(* IEC 61131-3 sources: CS_4_Aufzugsteuerung/src/Stations/CP112/Steuerung/Network, 1 file *)

(* ---- ConfigObjects.st ---- *)
FUNCTION GLOBAL TAB TASK_CONF
_K_TASK, _K_REAL,
_K_END_VAR,

_K_TASK, _K_CYCLIC,
_K_END_VAR,

_K_TASK, _K_BACKGROUND,
_K_END_VAR,

_K_END_CONF
END_FUNCTION

FUNCTION GLOBAL TAB IPR_CONF
_K_IPR
	0$UINT,
_K_END_VAR,
_K_END_CONF
END_FUNCTION

FUNCTION GLOBAL TAB CONFIG_TABLES
00096$UINT,
0$UINT, 1, 58, "_AXISBASE",
0$UINT, 1, 15, "_BUSINTERFACESDIASDRIVEMNG",
0$UINT, 0, 5, "_CAN",
0$UINT, 1, 11, "_CANLIB",
0$UINT, 1, 72, "_DRIVEAXIS",
0$UINT, 1, 81, "_DRIVEAXISBASE",
0$UINT, 1, 22, "_DRIVEAXISSET",
0$UINT, 1, 88, "_DRIVEMNG_DC062",
0$UINT, 1, 66, "_DRIVEMNGBASE",
0$UINT, 1, 20, "_FILESYS",
0$UINT, 0, 5, "_LINKER",
0$UINT, 1, 0, "_LMCABSENCODER",
0$UINT, 1, 117, "_LMCAXIS",
0$UINT, 2, 108, "_LMCAXISBASE",
0$UINT, 1, 32, "_LMCAXISREF",
0$UINT, 1, 41, "_LMCAXISVIS",
0$UINT, 1, 63, "_LMCAXISVISINT",
0$UINT, 1, 0, "_LMCAXISVISLOGHANDLE",
0$UINT, 1, 0, "_LMCAXISVISLOGVIEWER",
0$UINT, 1, 13, "_LMCAXISVISPARA",
0$UINT, 1, 1, "_LMCAXISVOVMONITORING",
0$UINT, 1, 75, "_LMCMATHFUNCTIONS",
0$UINT, 1, 1, "_LMCMODULEBASE",
0$UINT, 1, 0, "_LMCPUBLISHER",
0$UINT, 1, 11, "_LMCREFBASE",
0$UINT, 1, 21, "_LMCSAFETY",
0$UINT, 1, 1, "_MULTITASK",
0$UINT, 0, 5, "_OSKERNEL",
0$UINT, 1, 36, "_SERLIB",
0$UINT, 2, 0, "_STDLIB",
0$UINT, 1, 1, "_TASKOBJECTCONTROL",
0$UINT, 1, 69, "_VARANDRIVEBASE",
0$UINT, 1, 20, "AI043",
0$UINT, 1, 21, "ASCII_BIN",
0$UINT, 1, 26, "BUSINTERFACESDIAS",
0$UINT, 2, 1, "BUSINTERFACESDIASINTERNAL",
0$UINT, 1, 75, "BUSINTERFACEVARAN",
0$UINT, 0, 0, "CLSANTRIEB",
0$UINT, 0, 0, "CLSAUFZUGMODUL",
0$UINT, 0, 0, "CLSCOUNTER",
0$UINT, 0, 0, "CLSEMGSTOP_1",
0$UINT, 0, 0, "CLSENABLEDRIVE",
0$UINT, 0, 0, "CLSETAGENSENSORIK",
0$UINT, 0, 0, "CLSHAUPTABLAUF",
0$UINT, 0, 0, "CLSHMI",
0$UINT, 0, 0, "CLSMOTORCONTROL",
0$UINT, 0, 0, "CLSSIMPLECOUNTER",
0$UINT, 0, 0, "CLSTIMER",
0$UINT, 0, 0, "CLSTUERSENSORIK",
0$UINT, 1, 46, "CONTROLLER",
0$UINT, 1, 1, "CP112_IOS",
0$UINT, 0, 4, "CRITICALSECTION",
0$UINT, 2, 33, "DIASMASTER",
0$UINT, 1, 83, "DIASMASTERC",
0$UINT, 2, 25, "DIASMASTERMAIN",
0$UINT, 1, 0, "DIASMASTERPOSTSCAN",
0$UINT, 1, 13, "DM081",
0$UINT, 1, 14, "DM161",
0$UINT, 1, 87, "DRIVEPOSCONTROL",
0$UINT, 1, 11, "EEPROM",
0$UINT, 1, 21, "HUB_BASE",
0$UINT, 2, 11, "HUB_BASE_ROOT",
0$UINT, 2, 36, "HWBASE",
0$UINT, 2, 56, "HWBASECDIAS",
0$UINT, 1, 0, "HWCLOGGING",
0$UINT, 5, 27, "HWCONTROL",
0$UINT, 1, 10, "HWCONTROLBASE",
0$UINT, 1, 0, "HWRTPOSTSCAN",
0$UINT, 1, 6, "I2CCDIAS",
0$UINT, 1, 22, "MERKEREX",
0$UINT, 1, 17, "RAMEX",
0$UINT, 1, 9, "RAMFILE",
0$UINT, 1, 39, "SAFETYBASEFSOE",
0$UINT, 3, 19, "SAFETYCDIAS_BASE",
0$UINT, 2, 30, "SAFETYMANAGER",
0$UINT, 1, 4, "SAFETYUDP",
0$UINT, 1, 50, "SCP111",
0$UINT, 1, 60, "SDIASBASE",
0$UINT, 1, 10, "SDIASHUBBASE",
0$UINT, 1, 99, "SDIASMANAGER",
0$UINT, 2, 8, "SDIASPLC",
0$UINT, 1, 10, "SDIASSAFETYBASE",
0$UINT, 1, 41, "SDIASSAFETYMANAGERFSOE",
0$UINT, 1, 12, "SDM081",
0$UINT, 0, 46, "SIGCLIB",
0$UINT, 1, 11, "STRING",
0$UINT, 1, 86, "STRINGINTERNAL",
0$UINT, 1, 21, "SYNCCALL",
0$UINT, 2, 21, "VARAN_BASE",
0$UINT, 3, 8, "VARANMANAGER",
0$UINT, 2, 8, "VARANMANAGER_1",
0$UINT, 1, 26, "VARANMANAGER_BASE",
0$UINT, 1, 104, "VI021",
0$UINT, 1, 3, "VIRTUALBASEINIT",
0$UINT, 2, 11, "WATCHDOGDIAS",
0$UINT, 1, 2, "XXXBASE_IOS",
ONE_CFG$UINT, 0, 0, "ONE_HW_Network0",
ONE_CFG$UINT, 0, 0, "ONE_Motion",
ONE_CFG$UINT, 0, 0, "ONE_NW1",
ONE_CFG$UINT, 0, 0, "ONE_RT_EMG",
TASK_CFG$UINT, 0, 0, "TASK_CONF",
IPR_CFG$UINT, 0, 0, "IPR_CONF",
PRJ_CFG$UINT, 0, 0, "Steuerung",
END_FUNCTION

#ifdef __LSLLDR_IOELEMENTS__
FUNCTION GLOBAL TAB _IO_ELEMENTS_TAB
0001$UINT, 0014$UINT,
"**IOCONN_EMPTY**", "_DriveMng_DC0621.CmdState",
"IO_Element0", "DM0811.Output1",
"IO_Element1", "SCP1111.QuitComError",
"IO_Element5", "DM0811.Output2",
"IO_Element6", "DM0811.Output3",
"IO_Element7", "DM0811.Output4",
"xI_Emg1_1", "SDM0811.Safe_Input1",
"xI_Emg1_2", "SDM0811.Safe_Input2",
"xI_EnMotoren", "DM0811.Input4",
"xI_Etage0", "DM1611.Input1",
"xI_Etage1", "DM1611.Input2",
"xI_Etage2", "DM1611.Input3",
"xI_Etage3", "DM1611.Input4",
"xI_Lichtschranke", "DM0811.Input1",
0018$UINT,
"**IOCONN_EMPTY**", "_DriveMng_DC0621_Axis1.DriveMng",
"**IOCONN_EMPTY**", "_DriveMng_DC0622_Axis1.DriveMng",
"**IOCONN_EMPTY**", "DrivePosControl1.cDriveAxis",
"**IOCONN_EMPTY**", "_LMCAxis1.ActPosition",
"**IOCONN_EMPTY**", "DrivePosControl2.cDriveAxis",
"**IOCONN_EMPTY**", "_LMCAxis2.ActPosition",
"IO_Element0", "clsEnableDrive1.cOut1",
"IO_Element5", "clsEnableDrive1.cOut2",
"IO_Element6", "clsEnableDrive1.cOut3",
"IO_Element7", "clsEnableDrive1.cOut4",
"xI_Emg1_1", "clsEmgStop_1.c1",
"xI_Emg1_2", "clsEmgStop_1.c2",
"xI_EnMotoren", "clsEnableDrive1.cIn1",
"xI_Etage0", "clsHMI1.cTaster1",
"xI_Etage1", "clsHMI1.cTaster2",
"xI_Etage2", "clsHMI1.cTaster3",
"xI_Etage3", "clsHMI1.cTaster4",
"xI_Lichtschranke", "clsHMI1.cLichtschranke",
END_FUNCTION
#endif //__LSLLDR_IOELEMENTS__

FUNCTION GLOBAL TAB CH_REDIRECT_EMB_TAB
0000$UINT,
00023$UINT,
"_BUSINTERFACESDIASDRIVEMNG;SERIALNO", "\SERIALNOSTR.DATA",
"_DRIVEMNG_DC062;FWDATETR", "\FWDATESTRING.DATA",
"_DRIVEMNG_DC062;FWDATE", "\FWDATESTRING.DATA",
"_DRIVEMNG_DC062;FWNUMSTR", "\FWNUMSTRING.DATA",
"_DRIVEMNG_DC062;FWVERSION", "\FWNUMSTRING.DATA",
"_VARANDRIVEBASE;SERIALNO", "\SERIALNOSTR.DATA",
"AI043;SERIALNO", "\SERIALNOSTR.DATA",
"BUSINTERFACESDIAS;SERIALNO", "\SERIALNOSTR.DATA",
"BUSINTERFACEVARAN;SERIALNO", "\SERIALNOSTR.DATA",
"DM081;SERIALNO", "\SERIALNOSTR.DATA",
"DM161;SERIALNO", "\SERIALNOSTR.DATA",
"HWBASECDIAS;SERIALNO", "\SERIALNOSTR.DATA",
"SAFETYCDIAS_BASE;SERIALNO", "\SERIALNOSTR.DATA",
"SCP111;DESIGNERPRJNAME", "\SDIASSAFETYMANAGERFSOE1\PROJECTNAMESTR.DATA",
"SCP111;DESIGNERPRJREV", "\SDIASSAFETYMANAGERFSOE1\PROJECTREVISIONSTR.DATA",
"SCP111;SERIALNO", "\SERIALNOSTR.DATA",
"SDIASBASE;SERIALNO", "\SERIALNOSTR.DATA",
"SDIASSAFETYBASE;SERIALNO", "\SERIALNOSTR.DATA",
"SDIASSAFETYMANAGERFSOE;DESIGNERPRJNAME", "\PROJECTNAMESTR.DATA",
"SDIASSAFETYMANAGERFSOE;DESIGNERPRJREV", "\PROJECTREVISIONSTR.DATA",
"SDM081;SERIALNO", "\SERIALNOSTR.DATA",
"VARAN_BASE;SERIALNO", "\SERIALNOSTR.DATA",
"VI021;SERIALNO", "\SERIALNOSTR.DATA",
END_FUNCTION
